(* IEC 61131-3 sources: Test-Git_ESME26/TestProgettoESME_26.fbsproj/TemplateFullProgrammingFramework_Migration.device.xml.v3^/Plc Logic.plclogic.xml.v3^/Application.application.xml.v3^/TemplateFullProgrammingFramework/Examples/ExampleDiagSources/FB_ExampleTreeDiagSource.fb.st^, 6 files *)

(* ---- CancelWriting.meth.st ---- *)
{attribute 'hide'}
METHOD CancelWriting : BOOL
VAR_INPUT
END_VAR

(* Deactivate writing if we are (for whatever reason) no longer adressed.
   May happen in case network connection with Diagnostics is disrupted or Source will be disabled *)

THIS^.diOldCmd			:= 0;
THIS^.diCmdExecState	:= 0;

(* ---- DiagQuit.meth.st ---- *)
{attribute 'hide'}
METHOD DiagQuit : BOOL
VAR_INPUT
END_VAR

IF THIS^.i_xEnable AND THIS^.q_xActive AND THIS^.q_etDiag <> GD.ET_Diag.Ok AND THIS^.diState = 0 THEN

	THIS^.rtrigDiagQuit(CLK := THIS^.i_xDiagQuit);
	IF THIS^.rtrigDiagQuit.Q THEN
		CancelWriting();

		THIS^.udiOwnSourceId	:= 0;

		THIS^.fbTreeWriter.FB_Init(bInitRetains := FALSE, bInCopyCode := FALSE);

		THIS^.q_xReady		:= TRUE;
		THIS^.q_etDiag		:= GD.ET_Diag.Ok;
		THIS^.q_etDiagExt	:= ET_DiagExt.WaitUntilDiagnosticsManagerReady;
		THIS^.q_sMsg		:= '';

		THIS^.diState := 10;
	END_IF

END_IF

(* ---- ExceptionDuringWriting.meth.st ---- *)
{attribute 'hide'}
METHOD ExceptionDuringWriting : BOOL
VAR_INPUT
END_VAR

(* exception during writing *)
CASE THIS^.etDiagExtTPL OF
	TPL.ET_DiagExt.TreeStartAlreadySuccessfullyCalled,		// FB_TreeWriter.TreeStart
	TPL.ET_DiagExt.FileIdNotSet,							// FB_TreeWriter.TreeStart
	TPL.ET_DiagExt.FileIdInvalid,							// FB_TreeWriter.TreeStart & FB_TreeWriter.NodeStart & FB_TreeWriter.Parameter & FB_TreeWriter.NodeEnd & FB_TreeWriter.TreeEnd
	TPL.ET_DiagExt.FileNotOpen,								// FB_TreeWriter.TreeStart & FB_TreeWriter.NodeStart & FB_TreeWriter.Parameter & FB_TreeWriter.NodeEnd & FB_TreeWriter.TreeEnd
	TPL.ET_DiagExt.UnexpectedFeedback,						// FB_TreeWriter.TreeStart & FB_TreeWriter.NodeStart & FB_TreeWriter.Parameter & FB_TreeWriter.NodeEnd & FB_TreeWriter.TreeEnd
	TPL.ET_DiagExt.TreeStartNotCalled,						// FB_TreeWriter.NodeStart
	TPL.ET_DiagExt.TreeStartNotSuccessfullyCalled,			// FB_TreeWriter.NodeStart
	TPL.ET_DiagExt.NoMoreNodeOpen,							// FB_TreeWriter.Parameter & FB_TreeWriter.NodeEnd
	TPL.ET_DiagExt.CallTreeStartFirst,						// FB_TreeWriter.TreeEnd
	TPL.ET_DiagExt.NodesStillOpen:							// FB_TreeWriter.TreeEnd

		SetDiagOutputs(	i_etDiag	:= GD.ET_Diag.UnexpectedProgramBehavior,
						i_etDiagExt	:= ET_DiagExt.UnexpectedFeedback,
						i_sMsg		:= SE_CTBX.FC_MultiConcat(	i_sString1	:= 'FB_TreeWriter: ',
															i_sString2	:= GD.FC_EtDiagToString(THIS^.etDiag),
															i_sString3	:= ' - ',
															i_sString4	:= TPL.FC_EtDiagExtToString(THIS^.etDiagExtTPL)));
	ELSE
		SetDiagOutputs(	i_etDiag	:= GD.ET_Diag.UnexpectedProgramBehavior,
						i_etDiagExt	:= ET_DiagExt.UnexpectedFeedback,
						i_sMsg		:= SE_CTBX.FC_MultiConcat(	i_sString1	:= 'FB_TreeWriter: ',
															i_sString2	:= GD.FC_EtDiagToString(THIS^.etDiag),
															i_sString3	:= ' - ',
															i_sString4	:= TPL.FC_EtDiagExtToString(THIS^.etDiagExtTPL)));
END_CASE

CancelWriting();

(* ---- SetDiagOutputs.meth.st ---- *)
{attribute 'hide'}
METHOD SetDiagOutputs : BOOL
VAR_INPUT
	i_etDiag		: GD.ET_Diag;
	i_etDiagExt		: ET_DiagExt;
	i_sMsg			: STRING[80];
END_VAR

IF THIS^.q_etDiag = GD.ET_Diag.Ok OR i_etDiagExt = ET_DiagExt.Disabled THEN

	IF i_etDiag <> GD.ET_Diag.Ok OR i_etDiagExt = ET_DiagExt.Disabled THEN

		IF i_etDiag <> GD.ET_Diag.Ok THEN
			THIS^.iq_stComStructure.iq_diCmd := -THIS^.iq_stComStructure.iq_diCmd;
		END_IF

		IF i_etDiagExt = ET_DiagExt.Disabled THEN
			THIS^.q_xActive := FALSE;

			CancelWriting();
		END_IF

		THIS^.q_xReady := FALSE;
		THIS^.diState := 0;
	END_IF

	THIS^.q_etDiag		:= i_etDiag;
	THIS^.q_etDiagExt	:= i_etDiagExt;
	THIS^.q_sMsg		:= i_sMsg;

END_IF

(* ---- WriteDiagDataControl.meth.st ---- *)
{attribute 'hide'}
METHOD WriteDiagDataControl : BOOL
VAR_INPUT
END_VAR

IF (THIS^.diOldCmd <> THIS^.iq_stComStructure.iq_diCmd AND THIS^.iq_stComStructure.iq_diCmd > 0) THEN

	THIS^.diOldCmd := THIS^.iq_stComStructure.iq_diCmd;

	(* new command, start execution *)
	CASE THIS^.iq_stComStructure.iq_diCmd OF

		1: (* write diag data to file *)
			IF (THIS^.iq_stComStructure.i_diFileId > 0) THEN

				SetDiagOutputs(	i_etDiag		:= GD.ET_Diag.Ok,
								i_etDiagExt		:= ET_DiagExt.WritingToFile,
								i_sMsg			:= '');

				THIS^.iq_stComStructure.q_lrProgress := 0.0;

				THIS^.fbTreeWriter.diFileId := THIS^.iq_stComStructure.i_diFileId;

				THIS^.diCmdExecState := 1; (* start writing to file *)
			ELSE
				(* invalid file id *)
				SetDiagOutputs(	i_etDiag		:= GD.ET_Diag.InputParameterInvalid,
								i_etDiagExt		:= ET_DiagExt.FileIdInvalid,
								i_sMsg			:= CONCAT('Invalid file Id iq_stComStructure.i_diFileId: ', TO_STRING(THIS^.iq_stComStructure.i_diFileId)));
			END_IF
		ELSE
			(* unkown cmd *)
			SetDiagOutputs(	i_etDiag		:= GD.ET_Diag.InputParameterInvalid,
							i_etDiagExt		:= ET_DiagExt.CmdUnknown,
							i_sMsg			:= CONCAT('Unknown command iq_stComStructure.diCmd: ', DINT_TO_STRING(THIS^.iq_stComStructure.iq_diCmd)));

			CancelWriting();
	END_CASE
END_IF

(* ---- WriteDiagDataToFile.meth.st ---- *)
{attribute 'hide'}
METHOD WriteDiagDataToFile : BOOL
VAR_INPUT
END_VAR

TPL.FC_CanContinueWriting(iq_stCanContinueWriting := THIS^.iq_stComStructure.iq_stCanContinueWriting); (* loop as long as we can continue to write *)

WHILE (THIS^.iq_stComStructure.iq_stCanContinueWriting.xCanContinue) DO

	CASE THIS^.diCmdExecState OF
		1:
			(* start writing *)
			THIS^.fbTreeWriter.TreeStart(	i_sName					:= THIS^.c_sName,
											i_sTypeName				:= THIS^.c_sTypeName,
											i_sTitleEnglish			:= 'Example data as tree',
											i_sTitleGerman			:= 'Beispieldaten als Baum',
											i_uiPrintRank			:= 14,
											i_sEmptyListTextEnglish	:= 'No data available to show',
											i_sEmptyListTextGerman	:= 'Keine Daten zum Anzeigen vorhanden',
											q_etDiag				=> THIS^.etDiag,
											q_etDiagExt				=> THIS^.etDiagExtTPL);

			IF THIS^.etDiag <> GD.ET_Diag.Ok THEN
				ExceptionDuringWriting();
				EXIT;
			END_IF

			FOR THIS^.uiLevelCounter := 1 TO THIS^.c_uiMaxLevel DO
				THIS^.auiNodeCounter[uiLevelCounter] := 1;
			END_FOR

			THIS^.uiNodeId := 1;

			THIS^.lrSumNodes := ((1 - EXPT(THIS^.uiMaxNodePerLevel, THIS^.c_uiMaxLevel + 1)) / (1 - THIS^.uiMaxNodePerLevel));

			THIS^.uiLevelCounter := 1; (* start loop at index 1 *)

			THIS^.diCmdExecState := THIS^.diCmdExecState + 1;
		2:
			IF (THIS^.auiNodeCounter[THIS^.uiLevelCounter] <= THIS^.uiMaxNodePerLevel) THEN
				(* don't need to go up again, can create more nodes on this level *)

				(* create another subnode and go down *)
				(* create another node *)
				THIS^.uiNodeId := 0;
				THIS^.auiNodeCounter[THIS^.uiLevelCounter] := THIS^.auiNodeCounter[THIS^.uiLevelCounter] + 1;

				FOR THIS^.uiTmp := 1 TO THIS^.uiLevelCounter DO
					THIS^.uiNodeId := THIS^.uiNodeId * 100 + (THIS^.auiNodeCounter[THIS^.uiTmp] - 1);
				END_FOR

				THIS^.fbTreeWriter.NodeStart(	i_sName		:= CONCAT('Knoten_', UINT_TO_STRING(uiNodeId)),
												q_etDiag	=> THIS^.etDiag,
												q_etDiagExt	=> THIS^.etDiagExtTPL);

				IF THIS^.etDiag <> GD.ET_Diag.Ok THEN
					ExceptionDuringWriting();
					EXIT;
				END_IF

					THIS^.fbTreeWriter.Parameter(	i_sName		:= 'something',
													i_sValue	:= LREAL_TO_STRING(UINT_TO_LREAL(uiLevelCounter * auiNodeCounter[uiLevelCounter]) / UINT_TO_LREAL(uiNodeId)),
													q_etDiag	=> THIS^.etDiag,
													q_etDiagExt	=> THIS^.etDiagExtTPL);

					IF THIS^.etDiag <> GD.ET_Diag.Ok THEN
						ExceptionDuringWriting();
						EXIT;
					END_IF

				THIS^.uiLevelCounter := THIS^.uiLevelCounter + 1;

				IF (THIS^.uiLevelCounter > THIS^.c_uiMaxLevel) THEN
					(* go up again *)
					THIS^.fbTreeWriter.NodeEnd(	q_etDiag	=> THIS^.etDiag,
												q_etDiagExt	=> THIS^.etDiagExtTPL);

					IF THIS^.etDiag <> GD.ET_Diag.Ok THEN
						ExceptionDuringWriting();
						EXIT;
					END_IF

					THIS^.uiLevelCounter := THIS^.uiLevelCounter - 1;
				END_IF
			ELSE
				(* go up again *)
				THIS^.fbTreeWriter.NodeEnd(	q_etDiag	=> THIS^.etDiag,
											q_etDiagExt	=> THIS^.etDiagExtTPL);

				IF THIS^.etDiag <> GD.ET_Diag.Ok THEN
					ExceptionDuringWriting();
					EXIT;
				END_IF

				THIS^.auiNodeCounter[THIS^.uiLevelCounter] := 1; (* reset node counter of level *)

				THIS^.uiLevelCounter := THIS^.uiLevelCounter - 1;
				IF (THIS^.uiLevelCounter <= 1) THEN
					(* loop over all nodes and levels done *)
					THIS^.diCmdExecState := THIS^.diCmdExecState + 1;
				END_IF
			END_IF

			THIS^.iq_stComStructure.q_lrProgress := UINT_TO_LREAL(THIS^.auiNodeCounter[1]) * LREAL#100.0 / MAX(THIS^.lrSumNodes,0.0001);

		3:
			THIS^.fbTreeWriter.TreeEnd(	q_etDiag	=> THIS^.etDiag,
										q_etDiagExt	=> THIS^.etDiagExtTPL);

			IF THIS^.etDiag <> GD.ET_Diag.Ok THEN
				ExceptionDuringWriting();
				EXIT;
			END_IF
			(* done *)

			(* signal command execution *)
			THIS^.iq_stComStructure.iq_diCmd := 0;

			SetDiagOutputs(	i_etDiag	:= GD.ET_Diag.Ok,
							i_etDiagExt	:= ET_DiagExt.DataSuccessfullyWritten,
							i_sMsg		:= '');

			THIS^.diCmdExecState := 0;
			EXIT; (* exit the while loop *)
	END_CASE

	(* check again whether we can continue writing *)
	TPL.FC_CanContinueWriting(iq_stCanContinueWriting := THIS^.iq_stComStructure.iq_stCanContinueWriting);
END_WHILE
